// TwinCAT 3 PLC project EventLoggerSample
// ProgramVersion: 3.1.4026.26
// libraries:
//   EventFramework, * (DM)
//   Tc2_Standard, * (Beckhoff Automation GmbH)
//   Tc2_System, * (Beckhoff Automation GmbH)
//   Tc3_EventLogger, * (Beckhoff Automation GmbH)
// project tree:
//   GVLs/ GVL_EventTexts.TcGVL
//   POUs/ FB_Motor.TcPOU, MAIN.TcPOU
//   / PlcTask.TcTTO
// real-time tasks:
//   TASK PlcTask: cycle T#10ms, priority 20, ADS port 350

CONFIGURATION EventLoggerSample
    RESOURCE PLC ON TwinCAT3
        TASK PlcTask(INTERVAL := T#10ms, PRIORITY := 20);
        PROGRAM MAIN WITH PlcTask : MAIN;
    END_RESOURCE
END_CONFIGURATION

// ---- GVLs/GVL_EventTexts.TcGVL
// The event text list - the ONLY place to edit when adding an event. The TMC never changes.
//   nId       unique, stable number (source info id, HMI filter, key for external/CSV texts)
//   asText    one text per E_Language; {0}..{9} are replaced by the arguments
{attribute 'qualified_only'}
VAR_GLOBAL CONSTANT
	MachineStarted			: ST_EventDefinition := (nId := 100, eSeverity := TcEventSeverity.Info,		asText := ['Machine {0} started by {1}']);
	MachineStopped			: ST_EventDefinition := (nId := 101, eSeverity := TcEventSeverity.Info,		asText := ['Machine {0} stopped']);
	MotorHighTemperature	: ST_EventDefinition := (nId := 200, eSeverity := TcEventSeverity.Warning,	asText := ['Motor {0}: temperature high ({1} degC, limit {2} degC)']);
	MotorOverTemperature : ST_EventDefinition := (nId := 201, eSeverity := TcEventSeverity.Error,
							asText := ['Motor {0}: over temperature ({1} degC, limit {2} degC)',      // English
									   'Motor {0}: Übertemperatur ({1} °C, Grenze {2} °C)']);         // German
	MotorOverCurrent		: ST_EventDefinition := (nId := 202, eSeverity := TcEventSeverity.Error,	asText := ['Motor {0}: over current ({1} A, limit {2} A)']);
	DoorOpen				: ST_EventDefinition := (nId := 300, eSeverity := TcEventSeverity.Critical,	bWithConfirmation := TRUE, asText := ['Safety door {0} open']);
	DebugTrace				: ST_EventDefinition := (nId := 900, eSeverity := TcEventSeverity.Verbose,	asText := ['Trace: {0}']);
END_VAR

// ---- POUs/MAIN.TcPOU
PROGRAM MAIN
VAR
	// Simulation inputs - change them online
	fConveyorTemperature	: LREAL := 40.0;
	fConveyorCurrent		: LREAL := 5.0;
	fPumpTemperature		: LREAL := 40.0;
	fPumpCurrent			: LREAL := 5.0;
	bDoorOpen				: BOOL;
	bConfirmDoor			: BOOL;
	bStart					: BOOL;
	bStop					: BOOL;
	bTrace					: BOOL;

	fbConveyor	: FB_Motor;
	fbPump		: FB_Motor;

	fbDoorOpen	: FB_CatalogAlarm(stDefinition := GVL_EventTexts.DoorOpen);
	fbStarted	: FB_CatalogMessage(stDefinition := GVL_EventTexts.MachineStarted);
	fbStopped	: FB_CatalogMessage(stDefinition := GVL_EventTexts.MachineStopped);
	fbTrace		: FB_CatalogMessage(stDefinition := GVL_EventTexts.DebugTrace);

	rtStart		: R_TRIG;
	rtStop		: R_TRIG;
	rtTrace		: R_TRIG;
	rtConfirm	: R_TRIG;
END_VAR

// Two motors raise the same generic TMC events (e.g. GenericEvents.Error) at the same time
fbConveyor(sName := 'Conveyor', fTemperature := fConveyorTemperature, fCurrent := fConveyorCurrent);
fbPump(sName := 'Pump', fTemperature := fPumpTemperature, fCurrent := fPumpCurrent);

// Alarm with confirmation (bWithConfirmation in the text list)
fbDoorOpen.Arguments.Clear().AddString('Front');
fbDoorOpen.SetActive(bDoorOpen);
rtConfirm(CLK := bConfirmDoor);
IF rtConfirm.Q THEN
	fbDoorOpen.Confirm();
END_IF

// Messages
rtStart(CLK := bStart);
IF rtStart.Q THEN
	fbStarted.Arguments.Clear().AddString('Line 1').AddString('Operator');
	fbStarted.Send();
END_IF

rtStop(CLK := bStop);
IF rtStop.Q THEN
	fbStopped.Arguments.Clear().AddString('Line 1');
	fbStopped.Send();
END_IF

rtTrace(CLK := bTrace);
IF rtTrace.Q THEN
	fbTrace.Arguments.Clear().AddString('Conveyor temperature').AddLReal(fConveyorTemperature, 2);
	fbTrace.Send();
END_IF

END_PROGRAM

// ---- POUs/FB_Motor.TcPOU
// Example machine component. Its alarms share TMC events with every other motor;
// they can be active simultaneously because each alarm has its own source info.
FUNCTION_BLOCK FB_Motor
VAR_INPUT
	sName			: STRING(40);
	fTemperature	: LREAL;
	fCurrent		: LREAL;
END_VAR
VAR
	fbHighTemperature	: FB_CatalogAlarm(stDefinition := GVL_EventTexts.MotorHighTemperature);
	fbOverTemperature	: FB_CatalogAlarm(stDefinition := GVL_EventTexts.MotorOverTemperature);
	fbOverCurrent		: FB_CatalogAlarm(stDefinition := GVL_EventTexts.MotorOverCurrent);
END_VAR
VAR CONSTANT
	cWarnTemperature	: LREAL := 70.0;
	cMaxTemperature		: LREAL := 85.0;
	cMaxCurrent			: LREAL := 12.0;
END_VAR

// Arguments are refreshed every cycle but only taken over when the alarm is raised.
fbHighTemperature.Arguments.Clear().AddString(sName).AddLReal(fTemperature, 1).AddLReal(cWarnTemperature, 0);
fbHighTemperature.SetActive(fTemperature > cWarnTemperature AND fTemperature <= cMaxTemperature);

fbOverTemperature.Arguments.Clear().AddString(sName).AddLReal(fTemperature, 1).AddLReal(cMaxTemperature, 0);
fbOverTemperature.SetActive(fTemperature > cMaxTemperature);

fbOverCurrent.Arguments.Clear().AddString(sName).AddLReal(fCurrent, 2).AddLReal(cMaxCurrent, 1);
fbOverCurrent.SetActive(fCurrent > cMaxCurrent);

END_FUNCTION_BLOCK
